ABB RAPID module: TgtProg.mod

MODULE MainModule

GLOBAL Proc main()
    tool03.x = 0.125
    tool03.y = -0.375
    tool03.z = 123.457
    tool03.q1 = 0.923042
    tool03.q2 = -0.384698
    tool03.q3 = -0.000000
    tool03.q4 = 0.000001
    tool03.x = 0.000
    tool03.y = 0.000
    tool03.z = 0.000
    tool03.q1 = 0.000000
    tool03.q2 = 0.000000
    tool03.q3 = 0.000000
    tool03.q4 = 1.000000
    tool03.x = 0.000
    tool03.y = 0.000
    tool03.z = 0.000
    tool03.q1 = 0.000000
    tool03.q2 = 0.000000
    tool03.q3 = 1.000000
    tool03.q4 = -0.000000
    tool03.x = 0.000
    tool03.y = 0.000
    tool03.z = 0.000
    tool03.q1 = 0.000000
    tool03.q2 = 1.000000
    tool03.q3 = 0.000000
    tool03.q4 = -0.000000
EndProc
EndModule
